(* Logix 5000 project; controller SEAS_475 vendor 1 type 14 code 77 rev 17.4; software revision 17.01 *)

TASK MainTask (continuous, watchdog 500 ms) : MainProgram

MODULES
   Controller : vendor 1 type 14 code 77 (CompactLogixL32EController 0, rev 17.4)
      LocalENB : 1769-L32E Ethernet Port (CompactLogixL32Ethernet 1, rev 17.2)
         robot : ETHERNET-MODULE (Ethernet 192.168.1.100, rev 1.1, Output RPI 10 ms)
              robot:I.DATA[0].7   // TP Enable
              robot:I.DATA[0].6   // At Perch
              robot:I.DATA[0].5   // Fault
              robot:I.DATA[0].4   // Motion Held
              robot:I.DATA[0].3   // Program Paused
              robot:I.DATA[0].2   // Program Running
              robot:I.DATA[0].1   // System Ready
              robot:I.DATA[0].0   // CMD Enabled
              robot:I.DATA[0].8   // Batt Alarm
              robot:I.DATA[0].9   // Busy
              robot:I.DATA[0].10   // ACK1/SNO1
              robot:I.DATA[0].11   // ACK2/SNO2
              robot:I.DATA[0].12   // ACK3/SNO3
              robot:I.DATA[0].13   // ACK4/SNO4
              robot:I.DATA[0].14   // ACK5/SNO5
              robot:I.DATA[0].15   // ACK6/SNO6
              robot:I.DATA[0].16   // ACK7/SNO7
              robot:I.DATA[0].17   // ACK8/SNO8
              robot:I.DATA[0].18   // SNACK
              robot:I.DATA[0].19   // RESERVED
              robot:I.DATA[0].20   // HOPEN
              robot:I.DATA[0].21   // HCLOSED
              robot:I.DATA[0].25   // Wait Before Start
              robot:I.DATA[0].26   // Trigger Wire
              robot:I.DATA[0].27   // Slide
              robot:I.DATA[0].22   // DOUT 23
              robot:I.DATA[0].23   // DOUT 24
              robot:I.DATA[0].24   // DOUT 25
              robot:I.DATA[0].28   // DOUT 29
              robot:I.DATA[0].29   // DOUT 30
              robot:I.DATA[0].30   // DOUT 31
              robot:I.DATA[0].31   // DOUT 32
              robot:I.DATA[1].0   // DOUT 33
              robot:I.DATA[1].1   // DOUT 34
              robot:I.DATA[1].2   // DOUT 35
              robot:I.DATA[1].3   // DOUT 36
              robot:I.DATA[1].4   // DOUT 37
              robot:I.DATA[1].5   // DOUT 38
              robot:I.DATA[1].6   // DOUT 39
              robot:I.DATA[1].7   // DOUT 40
              robot:I.DATA[1].8   // DOUT 41
              robot:I.DATA[1].9   // DOUT 42
              robot:I.DATA[1].10   // DOUT 43
              robot:I.DATA[1].11   // DOUT 44
              robot:I.DATA[1].12   // DOUT 45
              robot:I.DATA[1].13   // DOUT 46
              robot:I.DATA[1].14   // DOUT 47
              robot:I.DATA[1].15   // DOUT 48
              robot:I.DATA[1].16   // DOUT 49
              robot:I.DATA[1].17   // DOUT 50
              robot:I.DATA[1].18   // DOUT 51
              robot:I.DATA[1].19   // DOUT 52
              robot:I.DATA[1].20   // DOUT 53
              robot:I.DATA[1].21   // DOUT 54
              robot:I.DATA[1].22   // DOUT 55
              robot:I.DATA[1].23   // DOUT 56
              robot:I.DATA[1].24   // DOUT 57
              robot:I.DATA[1].25   // DOUT 58
              robot:I.DATA[1].26   // DOUT 59
              robot:I.DATA[1].27   // DOUT 60
              robot:I.DATA[1].28   // DOUT 61
              robot:I.DATA[1].29   // DOUT 62
              robot:I.DATA[1].30   // DOUT 63
              robot:I.DATA[1].31   // DOUT 64
              robot:I.DATA[2].0   // DOUT 65
              robot:I.DATA[2].1   // DOUT 66
              robot:I.DATA[2].2   // DOUT 67
              robot:I.DATA[2].3   // DOUT 68
              robot:I.DATA[2].4   // DOUT 69
              robot:I.DATA[2].5   // DOUT 70
              robot:I.DATA[2].6   // DOUT 71
              robot:I.DATA[2].7   // DOUT 72
              robot:I.DATA[2].8   // DOUT 73
              robot:I.DATA[2].9   // DOUT 74
              robot:I.DATA[2].10   // DOUT 75
              robot:I.DATA[2].11   // DOUT 76
              robot:I.DATA[2].12   // DOUT 77
              robot:I.DATA[2].13   // DOUT 78
              robot:I.DATA[2].14   // DOUT 79
              robot:I.DATA[2].15   // DOUT 80
              robot:I.DATA[2].16   // DOUT 81
              robot:I.DATA[2].17   // SOUT 82
              robot:I.DATA[2].18   // DOUT 83
              robot:I.DATA[2].19   // DOUT 84
              robot:I.DATA[2].20   // DOUT 85
              robot:I.DATA[2].21   // DOUT 86
              robot:I.DATA[2].22   // DOUT 87
              robot:I.DATA[2].23   // DOUT 88
              robot:I.DATA[2].24   // DOUT 89
              robot:I.DATA[2].25   // DOUT 90
              robot:I.DATA[2].26   // DOUT 91
              robot:I.DATA[2].27   // DOUT 92
              robot:I.DATA[2].28   // DOUT 93
              robot:I.DATA[2].29   // DOUT 94
              robot:I.DATA[2].30   // DOUT 95
              robot:I.DATA[2].31   // DOUT 96
              robot:I.DATA[3].0   // DOUT 97
              robot:I.DATA[3].1   // DOUT 98
              robot:I.DATA[3].2   // DOUT 99
              robot:I.DATA[3].3   // DOUT 100
              robot:I.DATA[3].4   // DOUT 101
              robot:I.DATA[3].5   // DOUT 102
              robot:I.DATA[3].6   // DOUT 103
              robot:I.DATA[3].7   // DOUT 104
              robot:I.DATA[3].8   // DOUT 105
              robot:I.DATA[3].9   // DOUT 106
              robot:I.DATA[3].10   // DOUT 107
              robot:I.DATA[3].11   // DOUT 108
              robot:I.DATA[3].12   // DOUT 109
              robot:I.DATA[3].13   // DOUT 110
              robot:I.DATA[3].14   // DOUT 111
              robot:I.DATA[3].15   // DOUT 112
              robot:I.DATA[3].16   // DOUT 113
              robot:I.DATA[3].17   // DOUT 114
              robot:I.DATA[3].18   // DOUT 115
              robot:I.DATA[3].19   // DOUT 116
              robot:I.DATA[3].20   // DOUT 117
              robot:I.DATA[3].21   // DOUT 118
              robot:I.DATA[3].22   // DOUT 119
              robot:I.DATA[3].23   // DOUT 120
              robot:I.DATA[3].24   // DOUT 121
              robot:I.DATA[3].25   // DOUT 122
              robot:I.DATA[3].26   // DOUT 123
              robot:I.DATA[3].27   // DOUT 124
              robot:I.DATA[3].28   // DOUT 125
              robot:I.DATA[3].29   // DOUT 126
              robot:I.DATA[3].30   // DOUT 127
              robot:I.DATA[3].31   // DOUT 128
              robot:O.DATA[0].0   // IMSTP
              robot:O.DATA[0].1   // HOLD
              robot:O.DATA[0].2   // SFSPD
              robot:O.DATA[0].3   // CYCLE STOP
              robot:O.DATA[0].4   // FAULT RESET
              robot:O.DATA[0].5   // START
              robot:O.DATA[0].6   // HOME
              robot:O.DATA[0].7   // ENABLE
              robot:O.DATA[2].7   // DIN 72
              robot:O.DATA[0].8   // RSR1/PNS1/STYLE1
              robot:O.DATA[0].9   // RSR2/PNS2/STYLE2
              robot:O.DATA[0].10   // RSR3/PNS3/STYLE3
              robot:O.DATA[0].11   // RSR4/PNS4/STYLE4
              robot:O.DATA[0].12   // RSR5/PNS5/STYLE5
              robot:O.DATA[0].13   // RSR6/PNS6/STYLE6
              robot:O.DATA[0].14   // RSR7/PNS7/STYLE7
              robot:O.DATA[0].15   // RSR8/PNS8/STYLE8
              robot:O.DATA[0].16   // PNS strobe
              robot:O.DATA[0].17   // Prod start
              robot:O.DATA[1].31   // DIN 64
              robot:O.DATA[1].0   // DIN 33
              robot:O.DATA[0].18   // Hand Open
              robot:O.DATA[0].19   // Hand Closed
              robot:O.DATA[0].20   // DIN 21
              robot:O.DATA[0].21   // DIN 22
              robot:O.DATA[0].22   // DIN 23
              robot:O.DATA[0].23   // DIN 24
              robot:O.DATA[0].24   // DIN 25
              robot:O.DATA[0].25   // DIN 26
              robot:O.DATA[0].26   // DIN 27
              robot:O.DATA[0].27   // DIN 28
              robot:O.DATA[0].28   // DIN 29
              robot:O.DATA[0].29   // DIN 30
              robot:O.DATA[0].30   // DIN 31
              robot:O.DATA[0].31   // DIN 32
              robot:O.DATA[1].1   // DIN 34
              robot:O.DATA[1].2   // DIN 35
              robot:O.DATA[1].3   // DIN 36
              robot:O.DATA[1].4   // DIN 37
              robot:O.DATA[1].5   // DIN 38
              robot:O.DATA[1].6   // DIN 39
              robot:O.DATA[1].7   // DIN 40
              robot:O.DATA[1].8   // DIN 41
              robot:O.DATA[1].9   // DIN 42
              robot:O.DATA[1].10   // DIN 42
              robot:O.DATA[1].11   // DIN 44
              robot:O.DATA[1].12   // DIN 45
              robot:O.DATA[1].13   // DIN 46
              robot:O.DATA[1].14   // DIN 47
              robot:O.DATA[1].15   // DIN 48
              robot:O.DATA[1].16   // DIN 49
              robot:O.DATA[1].17   // DIN 50
              robot:O.DATA[1].18   // DIN 51
              robot:O.DATA[1].19   // DIN 52
              robot:O.DATA[1].20   // DIN 53
              robot:O.DATA[1].21   // DIN 54
              robot:O.DATA[1].22   // DIN 55
              robot:O.DATA[1].23   // DIN 56
              robot:O.DATA[1].24   // DIN 57
              robot:O.DATA[1].25   // DIN 58
              robot:O.DATA[1].26   // DIN 59
              robot:O.DATA[1].27   // DIN 60
              robot:O.DATA[1].28   // DIN 61
              robot:O.DATA[1].29   // DIN 62
              robot:O.DATA[1].30   // DIN 63
              robot:O.DATA[2].0   // DIN 65
              robot:O.DATA[2].1   // DIN 66
              robot:O.DATA[2].2   // DIN 67
              robot:O.DATA[2].3   // DIN 68
              robot:O.DATA[2].4   // DIN 69
              robot:O.DATA[2].5   // DIN 70
              robot:O.DATA[2].6   // DIN 71
              robot:O.DATA[2].8   // DIN 73
              robot:O.DATA[2].9   // DIN 74
              robot:O.DATA[2].10   // DIN 75
              robot:O.DATA[2].11   // DIN 76
              robot:O.DATA[2].12   // DIN 77
              robot:O.DATA[2].13   // DIN 78
              robot:O.DATA[2].14   // DIN 79
              robot:O.DATA[2].15   // DIN 80
              robot:O.DATA[2].16   // DIN 81
              robot:O.DATA[2].17   // DIN 82
              robot:O.DATA[2].18   // DIN 83
              robot:O.DATA[2].19   // DIN 84
              robot:O.DATA[2].20   // DIN 85
              robot:O.DATA[2].21   // DIN 86
              robot:O.DATA[2].22   // DIN 87
              robot:O.DATA[2].23   // DIN 88
              robot:O.DATA[2].24   // DIN 89
              robot:O.DATA[2].25   // DIN 90
              robot:O.DATA[2].26   // DIN 91
              robot:O.DATA[2].27   // DIN 92
              robot:O.DATA[2].28   // DIN 93
              robot:O.DATA[2].29   // DIN 94
              robot:O.DATA[2].30   // DIN 95
              robot:O.DATA[2].31   // DIN 96
              robot:O.DATA[3].0   // DIN 97
              robot:O.DATA[3].1   // DIN 98
              robot:O.DATA[3].2   // DIN 99
              robot:O.DATA[3].3   // DIN 100
              robot:O.DATA[3].4   // DIN 101
              robot:O.DATA[3].5   // DIN 102
              robot:O.DATA[3].6   // DIN 103
              robot:O.DATA[3].7   // DIN 104
              robot:O.DATA[3].8   // DIN 105
              robot:O.DATA[3].9   // DIN 106
              robot:O.DATA[3].10   // DIN 107
              robot:O.DATA[3].11   // DIN 108
              robot:O.DATA[3].12   // DIN 109
              robot:O.DATA[3].13   // DIN 110
              robot:O.DATA[3].14   // DIN 111
              robot:O.DATA[3].15   // DIN 112
              robot:O.DATA[3].16   // DIN 113
              robot:O.DATA[3].17   // DIN 114
              robot:O.DATA[3].18   // DIN 115
              robot:O.DATA[3].19   // DIN 116
              robot:O.DATA[3].20   // DIN 117
              robot:O.DATA[3].21   // DIN 118
              robot:O.DATA[3].22   // DIN 119
              robot:O.DATA[3].23   // DIN 120
              robot:O.DATA[3].24   // DIN 121
              robot:O.DATA[3].25   // DIN 122
              robot:O.DATA[3].26   // DIN 123
              robot:O.DATA[3].27   // DIN 124
              robot:O.DATA[3].28   // DIN 125
              robot:O.DATA[3].29   // DIN 126
              robot:O.DATA[3].30   // DIN 127
              robot:O.DATA[3].31   // DIN 128
      Local : CompactBus (CompactVirtualAdapter 3, rev 17.2, Input RPI 5 ms)
         Input_2 : 1769-IQ16 (Compact 2, rev 1.1, Input RPI 5 ms)
              Local:2:I.DATA.0   // Start Button
              Local:2:I.DATA.1   // Stop Button (paused)
              Local:2:I.DATA.2   // Reset Button
              Local:2:I.DATA.3   // Push Button 1 (Restart)
              Local:2:I.DATA.4   // Push Button 2
              Local:2:I.DATA.5   // Push Button 3
              Local:2:I.DATA.6   // Key Switch
              Local:2:I.DATA.7   // Selector Switch
              Local:2:I.DATA.8   // Robot input 1
              Local:2:I.DATA.9   // robot input 2
              Local:2:I.DATA.10   // robot input 3
              Local:2:I.DATA.11   // robot input 4
              Local:2:I.DATA.12   // robot input 5
              Local:2:I.DATA.13   // robot input 6
              Local:2:I.DATA.14   // Open
              Local:2:I.DATA.15   // Open
         Input_Output2 : vendor 1 type 7 code 66 (Compact 5, rev 2.1, Output RPI 5 ms)
              Local:5:I.DATA.0   // Open
              Local:5:I.DATA.1   // Open
              Local:5:I.DATA.2   // Open
              Local:5:I.DATA.3   // Open
              Local:5:I.DATA.4   // Open
              Local:5:I.DATA.5   // Open
              Local:5:O.DATA.0   // Camera Trigger
              Local:5:O.DATA.1   // Open
              Local:5:O.DATA.2   // Open
              Local:5:O.DATA.3   // Open
         Input_Output1 : vendor 1 type 7 code 66 (Compact 4, rev 2.1, Output RPI 5 ms)
              Local:4:I.DATA.0   // Open
              Local:4:I.DATA.1   // Open
              Local:4:I.DATA.2   // Open
              Local:4:I.DATA.3   // Open
              Local:4:I.DATA.4   // Open
              Local:4:I.DATA.5   // Open
              Local:4:O.DATA.0   // Light Tree Red
              Local:4:O.DATA.1   // Light Tree Yellow
              Local:4:O.DATA.2   // Light Tree Green
              Local:4:O.DATA.3   // Light Tree Blue
         Input_1 : 1769-IQ16 (Compact 1, rev 1.1, Input RPI 5 ms)
              Local:1:I.DATA.0   // Front Panel Start
              Local:1:I.DATA.1   // Front Panel Stop
              Local:1:I.DATA.2   // Front Panel Key Switch
              Local:1:I.DATA.3   // Front Panel Reset
              Local:1:I.DATA.4   // Red PB1
              Local:1:I.DATA.5   // Red PB2
              Local:1:I.DATA.6   // Red PB3
              Local:1:I.DATA.7   // Red PB4
              Local:1:I.DATA.8   // Open
              Local:1:I.DATA.9   // Open
              Local:1:I.DATA.10   // Open
              Local:1:I.DATA.11   // Open
              Local:1:I.DATA.12   // Open
              Local:1:I.DATA.13   // Open
              Local:1:I.DATA.14   // Open
              Local:1:I.DATA.15   // Open
         Output_1 : 1769-OB16 (Compact 3, rev 2.1, Output RPI 5 ms)
              Local:3:O.DATA.0   // Start Light
              Local:3:O.DATA.1   // Reset Light
              Local:3:O.DATA.2   // Push Button 1 Light
              Local:3:O.DATA.3   // Push Button 2 Light
              Local:3:O.DATA.4   // Push Button 3 Light
              Local:3:O.DATA.5   // Indicator Light 1
              Local:3:O.DATA.6   // Indicator Light 2
              Local:3:O.DATA.8   // Robot Hand Open
              Local:3:O.DATA.9   // Robot Hand Closed
              Local:3:O.DATA.7   // Audio Alarm
              Local:3:O.DATA.10   // Slide On
         Output_2 : 1769-OB16 (Compact 6, rev 2.1, Output RPI 5 ms)
              Local:6:O.DATA.1   // Front Panel Reset Light
              Local:6:O.DATA.0   // Front Panel Start Light
              Local:6:O.DATA.2   // Front Panel Q1 Light
              Local:6:O.DATA.3   // Front Panel Q2 Light
              Local:6:O.DATA.4   // Open
              Local:6:O.DATA.5   // Open
              Local:6:O.DATA.6   // Open
              Local:6:O.DATA.7   // Open
END_MODULES

VAR_GLOBAL   (* controller tags *)
   b1 : DINT;
   B2 : DINT;
        .0   // Start over bit
   B3_10_Fanuc_Produced_DIN_3 : DINT; {produced}
        .0   // DIN 65
        .1   // DIN 66
        .2   // DIN 67
        .3   // DIN 68
        .4   // DIN 69
        .5   // DIN 70
        .6   // DIN 71
        .7   // DIN 72
        .8   // DIN 73
        .9   // DIN 74
        .10   // DIN 75
        .11   // DIN 76
        .12   // DIN 77
        .13   // DIN 78
        .14   // DIN 79
        .15   // DIN 80
        .16   // DIN 81
        .17   // DIN 82
        .18   // DIN 83
        .19   // DIN 84
        .20   // DIN 85
        .21   // DIN 86
        .22   // DIN 87
        .23   // DIN 88
        .24   // DIN 89
        .25   // DIN 90
        .26   // DIN 91
        .27   // DIN 92
        .28   // DIN 93
        .29   // DIN 94
        .30   // DIN 95
        .31   // DIN 96
   B3_11_Fanuc_Produced_DOUT_3 : DINT; {produced}
        .0   // DOUT 65
        .1   // DOUT 66
        .2   // DOUT 67
        .3   // DOUT 68
        .4   // DOUT 69
        .5   // DOUT 70
        .6   // DOUT 71
        .7   // DOUT 72
        .8   // DOUT 73
        .9   // DOUT 74
        .10   // DOUT 75
        .11   // DOUT 76
        .12   // DOUT 77
        .13   // DOUT 78
        .14   // DOUT 79
        .15   // DOUT 80
        .16   // DOUT 81
        .17   // DOUT 82
        .18   // DOUT 83
        .19   // DOUT 84
        .20   // DOUT 85
        .21   // DOUT 86
        .22   // DOUT 87
        .23   // DOUT 88
        .24   // DOUT 89
        .25   // DOUT 90
        .26   // DOUT 91
        .27   // DOUT 92
        .28   // DOUT 93
        .29   // DOUT 94
        .30   // DOUT 95
        .31   // DOUT 96
   B3_12_Fanuc_Produced_DIN_4 : DINT; {produced}
        .0   // DIN 97
        .1   // DIN 98
        .2   // DIN 99
        .3   // DIN 100
        .4   // DIN 101
        .5   // DIN 102
        .6   // DIN 103
        .7   // DIN 104
        .8   // DIN 105
        .9   // DIN 106
        .10   // DIN 107
        .11   // DIN 108
        .12   // DIN 109
        .13   // DIN 110
        .14   // DIN 111
        .15   // DIN 112
        .16   // DIN 113
        .17   // DIN 114
        .18   // DIN 115
        .19   // DIN 116
        .20   // DIN 117
        .21   // DIN 118
        .22   // DIN 119
        .23   // DIN 120
        .24   // DIN 121
        .25   // DIN 122
        .26   // DIN 123
        .27   // DIN 124
        .28   // DIN 125
        .29   // DIN 126
        .30   // DIN 127
        .31   // DIN 128
   B3_13_Fanuc_Produced_DOUT_4 : DINT; {produced}
        .0   // DOUT 97
        .1   // DOUT 98
        .2   // DOUT 99
        .3   // DOUT 100
        .4   // DOUT 101
        .5   // DOUT 102
        .6   // DOUT 103
        .7   // DOUT 104
        .8   // DOUT 105
        .9   // DOUT 106
        .10   // DOUT 107
        .11   // DOUT 108
        .12   // DOUT 109
        .13   // DOUT 110
        .14   // DOUT 111
        .15   // DOUT 112
        .16   // DOUT 113
        .17   // DOUT 114
        .18   // DOUT 115
        .19   // DOUT 116
        .20   // DOUT 117
        .21   // DOUT 118
        .22   // DOUT 119
        .23   // DOUT 120
        .24   // DOUT 121
        .25   // DOUT 122
        .26   // DOUT 123
        .27   // DOUT 124
        .28   // DOUT 125
        .29   // DOUT 126
        .30   // DOUT 127
        .31   // DOUT 128
   B3_2_L32_Produced_Outputs_1 : DINT := 327682; {produced}
        .0   // Start Light
        .1   // Reset Light
        .7   // Audio Alarm
        .10   // Slide On
        .11   // Open
        .12   // Open
        .13   // Open
        .14   // Open
        .15   // Open
        .21   // Open
        .22   // Open
        .23   // Open
        .28   // Open
        .29   // Open
        .30   // Open
        .31   // Open
        .2   // Push Button 1 Light
        .3   // Push Button 2 Light
        .4   // Push Button 3 Light
        .5   // Indicator Light 1
        .6   // Indicator Light 2
        .8   // Robot Hand Open
        .9   // Robot Hand Close
        .16   // Light Tree Red
        .17   // Light Tree Yellow
        .18   // Light Tree Green
        .19   // Light Tree Blue
        .20   // Camera Trigger
        .24   // Front Panel Start Light
        .25   // Front Panel Reset Light
        .26   // Front Panel Q1 Light
        .27   // Front Panel Q2 Light
   B3_3_L32_Produced_Inputs_1 : DINT := 131074; {produced}
        .4   // Reb PB1
        .5   // Red PB2
        .6   // Red PB3
        .7   // Red PB4
        .9   // Open
        .10   // Open
        .11   // Open
        .12   // Open
        .13   // Open
        .14   // Open
        .15   // Open
        .16   // Start Button
        .18   // Reset Button
        .22   // Key Switch
        .30   // Open
        .31   // Open
        .8   // Open
        .0   // Front Panel Start
        .1   // Front Panel Stop
        .2   // Front Panel Key
        .3   // Front Panel Reset
        .17   // Stop Button (Pause)
        .19   // Push Button 1 (restart)
        .20   // Push Button 2
        .21   // Push Button 3
        .23   // Selector Switch
        .24   // Robot Input 1
        .25   // Robot Input 2
        .26   // Robot Input 3
        .27   // Robot Input 4
        .28   // Robout Input 5
        .29   // Robout Input 6
   B3_4_L32_Produced_Output_2 : DINT; {produced}
        .1   // Not Wired
        .2   // Not Wired
        .3   // Not Wired
        .4   // Not Wired
        .5   // Not Wired
        .6   // Not Wired
        .7   // Not Wired
        .0   // Not Wired
   B3_5_L32_Produced_Inputs_2 : DINT; {produced}
        .0   // Open
        .1   // Open
        .2   // Open
        .3   // Open
        .4   // Open
        .5   // Open
        .6   // Open
        .7   // Open
        .8   // Open
        .9   // Open
        .10   // Open
        .11   // Open
   B3_6_Fanuc_Produced_DIN_1 : DINT := 135; {produced}
        .0   // *IMSTP
        .1   // *HOLD
        .2   // *SFSPD
        .3   // CYCLE STOP
        .4   // FAULT RESSET
        .5   // START
        .7   // ENABLE
        .16   // PNS Strobe
        .17   // Prod Start
        .18   // Hand Open
        .19   // Hand Closed
        .20   // DIN 21
        .21   // DIN 22
        .22   // DIN 23
        .23   // DIN 24
        .24   // DIN 25
        .25   // DIN 26
        .26   // DIN 27
        .27   // DIN 28
        .28   // DIN 29
        .29   // DIN 30
        .30   // DIN 31
        .31   // DIN 32
        .6   // HOME
        .8   // RSR1/PNS1/STYLE1
        .9   // RSR2/PNS2/STYLE2
        .10   // RSR3/PNS3/STYLE3
        .11   // RSR4/PNS4/STYLE4
        .12   // RSR5/PNS5/STYLE5
        .13   // RSR6/PNS6/STYLE6
        .14   // RSR7/PNS7/STYLE7
        .15   // RSR8/PNS8/STYLE8
   B3_7_Fanuc_Produced_DOUT_1 : DINT := 160; {produced}
        .0   // CMD Enabled
        .1   // System Ready
        .2   // PRG running
        .3   // Prg Paused
        .4   // Motion held
        .5   // Fault
        .6   // At perch
        .7   // TP Enabled
        .8   // Battery Alarm
        .9   // Busy
        .10   // ACK1/SNO1
        .11   // ACK2/SNO2
        .12   // ACK3/SNO3
        .13   // ACK4/SNO4
        .14   // ACK5/SNO5
        .15   // ACK6/SNO6
        .16   // ACK7/SNO7
        .18   // SNACK
        .20   // HOEPN
        .21   // HCLOSED
        .22   // DOUT 23
        .23   // DOUT 24
        .31   // DOUT 32
        .30   // DOUT 31
        .27   // Slide
        .28   // DOUT 29
        .29   // DOUT 30
        .24   // DOUT 25
        .19   // Reserved
        .26   // Trigger Wire
        .25   // Wait Before Start
        .17   // ACK8/SNO8
   B3_8_Fanuc_Produced_DIN_2 : DINT; {produced}
        .11   // DIN 44
        .12   // DIN 45
        .13   // DIN 46
        .14   // DIN 47
        .15   // DIN 48
        .16   // DIN 49
        .17   // DIN 50
        .18   // DIN 51
        .19   // DIN 52
        .20   // DIN 53
        .21   // DIN 54
        .22   // DIN 55
        .23   // DIN 56
        .24   // DIN 57
        .25   // DIN 58
        .26   // DIN 59
        .27   // DIN 60
        .28   // DIN 61
        .29   // DIN 62
        .30   // DIN 63
        .31   // DIN 64
        .0   // DIN 33
        .1   // DIN 34
        .2   // DIN 35
        .3   // DIN 36
        .4   // DIN 37
        .5   // DIN 38
        .6   // DIN 39
        .7   // DIN 40
        .8   // DIN 41
        .9   // DIN 42
        .10   // DIN 43
   B3_9_Fanuc_Produced_DOUT_2 : DINT; {produced}
        .0   // DOUT 33
        .1   // DOUT 34
        .2   // DOUT 35
        .3   // DOUT 36
        .4   // DOUT 37
        .5   // DOUT 38
        .6   // DOUT 39
        .7   // DOUT 40
        .8   // DOUT 41
        .9   // DOUT 42
        .10   // DOUT 43
        .11   // DOUT 44
        .12   // DOUT 45
        .13   // DOUT 46
        .14   // DOUT 47
        .15   // DOUT 48
        .16   // DOUT 49
        .17   // DOUT 50
        .18   // DOUT 51
        .19   // DOUT 52
        .20   // DOUT 53
        .21   // DOUT 54
        .22   // DOUT 55
        .23   // DOUT 56
        .24   // DOUT 57
        .25   // DOUT 58
        .26   // DOUT 59
        .27   // DOUT 60
        .28   // DOUT 61
        .29   // DOUT 62
        .30   // DOUT 63
        .31   // DOUT 64
   C1 : COUNTER := (PRE := 1, ACC := 5, CU := 1, DN := 1);   // Stop button counter
   C2 : COUNTER := (PRE := 4, ACC := 21, DN := 1);   // Reset light counter
   Pause_Bit : DINT;
   push_button_1_timer : TIMER := (PRE := 10000, ACC := 10000, EN := 1, DN := 1);
   PUSH_BUTTON_BITS : DINT;
   t1 : TIMER := (PRE := 300);   // pulse timer
   t2 : TIMER := (PRE := 100);   // on
   t3 : TIMER := (PRE := 200);   // off
   t4 : TIMER := (PRE := 300);
END_VAR

PROGRAM MainProgram   (* main routine MainRoutine *)
VAR
   Fanuc_Invis : BOOL;
   Fanuc_Mov : COUNTER := (PRE := 1, ACC := 1, DN := 1);
   Fanuc_Mov_Cam1 : TIMER := (PRE := 40000, ACC := 40000, EN := 1, DN := 1);
   Fanuc_Mov_Perch : TIMER := (PRE := 27000, ACC := 27000, EN := 1, DN := 1);
   Fanuc_mov_Steve : TIMER := (PRE := 40000);
   Fanuc_Rot_invs : BOOL := 1;
   Fanuc_Stationary : BOOL;
   HMI_Reset_Light : BOOL := 1;
   Reset_for_HMI : BOOL;
   Start_for_HMI : BOOL;
   steve_arm1_invis : BOOL := 1;
   steve_arm2_invis : BOOL := 1;
   steve_mov_bk : TIMER := (PRE := 25000, ACC := 25000, EN := 1, DN := 1);
   Steve_Move_Timer : TIMER := (PRE := 15000, ACC := 15000, EN := 1, DN := 1);
   Steve_perch : BOOL;
   Stop_for_HMI : BOOL;
   System_Ready_HMI : BOOL;
END_VAR

ROUTINE MainRoutine   (* ladder *)
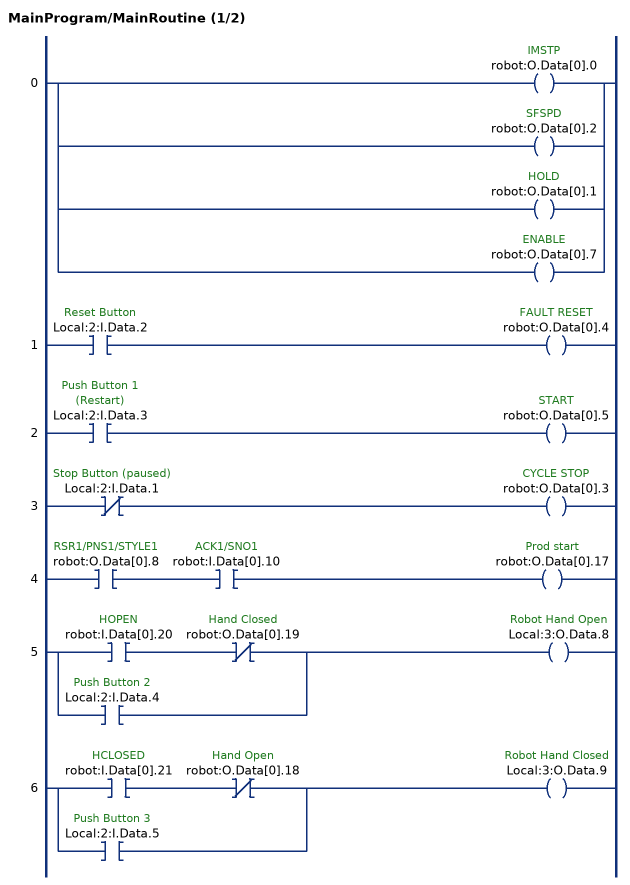
   0: [OTE(robot:O.Data[0].0) ,[OTE(robot:O.Data[0].2) ,[OTE(robot:O.Data[0].1) ,OTE(robot:O.Data[0].7) ] ] ];
   1: XIC(Local:2:I.Data.2)OTE(robot:O.Data[0].4);
   2: XIC(Local:2:I.Data.3)OTE(robot:O.Data[0].5);
   3: XIO(Local:2:I.Data.1)OTE(robot:O.Data[0].3);
   4: XIC(robot:O.Data[0].8)XIC(robot:I.Data[0].10)OTE(robot:O.Data[0].17);
   5: [XIC(robot:I.Data[0].20) XIO(robot:O.Data[0].19) ,XIC(Local:2:I.Data.4) ]OTE(Local:3:O.Data.8);
   6: [XIC(robot:I.Data[0].21) XIO(robot:O.Data[0].18) ,XIC(Local:2:I.Data.5) ]OTE(Local:3:O.Data.9);
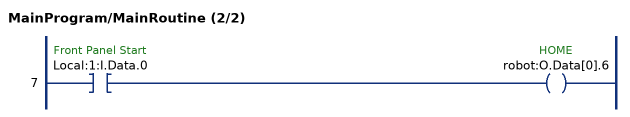
   7: XIC(Local:1:I.Data.0)OTE(robot:O.Data[0].6);
END_ROUTINE
END_PROGRAM
